// TIA Portal V21 export
// export: Created 2026-11-10T07:35:03.4177775Z, ExportSetting WithDefaults, DisplayName Totally Integrated Automation Portal, DisplayVersion V21 Update 3, DisplayName STEP 7 Professional, DisplayVersion V21 Update 3, DisplayName STEP 7 Safety, DisplayVersion V21, DisplayName Tech WebApplication, DisplayVersion V21, DisplayName WinCC Basic/Comfort/Advanced, DisplayVersion V21 Update 3, DisplayName WinCC Unified, DisplayVersion V21 Update 3
FUNCTION_BLOCK "FB_Lad_ex036"   // FB66, LAD
{ S7_Optimized_Access := 'TRUE' }
VERSION : 0.1
// stored: AutoNumber true, IsIECCheckEnabled false, IsRetainMemResEnabled false, MemoryReserve 100, SetENOAutomatically false, UDAEnableTagReadback false
   VAR_INPUT
      v_size : DInt;
      v_out : WString;
   END_VAR
   VAR_IN_OUT
      v_variable : Array[0..99] of Byte;
   END_VAR
BEGIN

REGION Network 1: GetSymbolName - Read out a tag on the input parameter
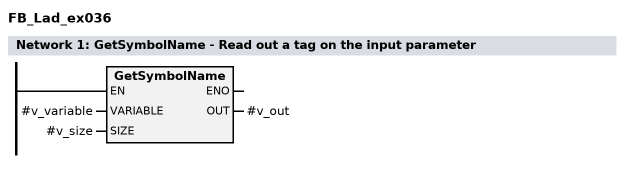
   RUNG wire#powerrail
      GetSymbolName(variable := #v_variable, size := #v_size, OUT => #v_out)
   END_RUNG
   // the same network as SCL:
   GetSymbolName(variable := #v_variable, size := #v_size, OUT => #v_out);
END_REGION
END_FUNCTION_BLOCK
